// TIA Portal V21 export
// export: Created 2026-11-10T19:11:41.9252955Z, ExportSetting WithDefaults, DisplayName Totally Integrated Automation Portal, DisplayVersion V21 Update 3, DisplayName STEP 7 Professional, DisplayVersion V21 Update 3, DisplayName STEP 7 Safety, DisplayVersion V21, DisplayName Tech WebApplication, DisplayVersion V21, DisplayName WinCC Basic/Comfort/Advanced, DisplayVersion V21 Update 3, DisplayName WinCC Unified, DisplayVersion V21 Update 3
DATA_BLOCK "DB_URCV_SFB"   // DB53
// stored: AutoNumber true, DBAccessibleFromOPCUA true, DBAccessibleFromWebserver true, InstanceOfName URCV_SFB, OfSystemLibElement URCV, OfSystemLibVersion 1.2
"URCV_SFB"
   // VAR_INPUT
   //    EN_R : Bool;
   //    ID : CONN_PRG;
   //    R_ID : CONN_R_ID;
   // END_VAR
   // VAR_OUTPUT
   //    NDR : Bool;
   //    ERROR : Bool;
   //    STATUS : Word;
   // END_VAR
   // VAR_IN_OUT
   //    RD_1 : Variant;
   //    RD_2 : Variant;
   //    RD_3 : Variant;
   //    RD_4 : Variant;
   // END_VAR
   // VAR
   //    INDEX : Word;
   // END_VAR
BEGIN
END_DATA_BLOCK
